(* IEC 61131-3 sources: plcassist-cli/packages/volt-lsp-iec/test-corpus/awa-palletizer/Device/Plc Logic/Application/Library Manager/L_SPMI_PlcParameterManager, 22 files *)

(* ---- L_SPMI_CONSTANT_DEFINES.gvl ---- *)
VAR_GLOBAL
	APPLICATION_AREA_0 : DINT := 0;
	APPLICATION_AREA_1 : DINT := 1;
	APPLICATION_AREA_2 : DINT := 2;
	APPLICATION_AREA_3 : DINT := 3;
END_VAR

(* ---- L_SPMI_LEM_ACCESS.gvl ---- *)
VAR_GLOBAL
	BASIC_SETTINGS : UINT := 4;
	REFID_PLCPM : UINT := 16#2801;
	EVTID_INF_INIT_WRITE : UINT := 16#1101;
	EVTID_INF_DEFAULT_WRITE : UINT := 16#1102;
	EVTID_WRN_INIT_PARAMETER : UINT := 16#1201;
	EVTID_WRN_LOAD_FACTORYSETTINGS : UINT := 16#1202;
	EVTID_WRN_LOAD_TADEFAULTS : UINT := 16#1203;
	EVTID_ERR_REGISTRATION : UINT := 16#1401;
	EVTID_ERR_OPEN_LXD_FILE : UINT := 16#1402;
	EVTID_ERR_OPEN_PRM_FILE : UINT := 16#1403;
	EVTPAR_DT_BOOL : INT := 1;
	EVTPAR_DT_S8 : INT := 2;
	EVTPAR_DT_S16 : INT := 3;
	EVTPAR_DT_S32 : INT := 4;
	EVTPAR_DT_U8 : INT := 5;
	EVTPAR_DT_U16 : INT := 6;
	EVTPAR_DT_U32 : INT := 7;
	EVTPAR_DT_STR_UNI_CODE8 : INT := 8;
	EVTPAR_DT_STR_ASCII : INT := 9;
	EVTPAR_DT_BYTE_ARRAY : INT := 10;
	EVTPAR_DT_S64 : INT := 11;
	EVTPAR_DT_U64 : INT := 12;
	EVTPAR_DT_FLOAT_32 : INT := 13;
	EVTPAR_DT_FLOAT_64 : INT := 14;
END_VAR

(* ---- L_SPMI_ITF_PLCPARAMETERMANAGER.itf ---- *)
INTERFACE L_SPMI_ITF_PLCPARAMETERMANAGER
END_INTERFACE

METHOD GETPARAMETEROBJECT : POINTER TO L_SPMI_ParameterObject
VAR_INPUT
	WINDEX : WORD;
	BYSUBINDEX : BYTE;
	PNUMSUBOBJECTS : POINTER TO BYTE;
END_VAR
END_METHOD

METHOD GETPARAMETEROBJECTLIST : L_SPMI_ParameterObjectList
END_METHOD

METHOD GETPARAMETERVALUE : RTS_IEC_RESULT
VAR_INPUT
	PARAMETERADDRESS : L_SPMI_ParameterAddress;
	PPARAMETERVALUE : POINTER TO L_SPMI_ParameterValueInfo;
END_VAR
END_METHOD

METHOD GETSUBOBJECTRECORDINFO : L_SPMI_SubObjectRecordInfo
VAR_INPUT
	WINDEX : WORD;
END_VAR
END_METHOD

METHOD LOADFACTORYSETTINGS : RTS_IEC_RESULT
END_METHOD

METHOD LOADPARAMETERSET : RTS_IEC_RESULT
END_METHOD

METHOD LOADTADEFAULTPARAMETER : RTS_IEC_RESULT
END_METHOD

METHOD RELAODPARAMETERDESCRIPTION : RTS_IEC_RESULT
END_METHOD

METHOD SAVEPARAMETERSET : RTS_IEC_RESULT
END_METHOD

METHOD SETPARAMETERVALUE : RTS_IEC_RESULT
VAR_INPUT
	PARAMETERADDRESS : L_SPMI_ParameterAddress;
	PPARAMETERVALUE : POINTER TO L_SPMI_ParameterValueInfo;
END_VAR
END_METHOD

METHOD UPDATEONLINECHANGEDPARAMETER : RTS_IEC_RESULT
END_METHOD

(* ---- L_SPMI_UTITF_PLCPM.itf ---- *)
INTERFACE L_SPMI_UTITF_PLCPM
END_INTERFACE

METHOD UT_WRITEPARAMETERVALUE : RTS_IEC_RESULT
VAR_INPUT
	PPARAMETEROBJECT : POINTER TO L_SPMI_ParameterObject;
	PPARAMETERVALUE : POINTER TO L_SPMI_ParameterValueInfo;
	BISDEFAULT : BOOL;
END_VAR
END_METHOD

(* ---- GETBOOLEANPROPERTY.fun ---- *)
FUNCTION GETBOOLEANPROPERTY : BOOL
VAR_INPUT
	STKEY : WSTRING;
END_VAR
END_FUNCTION

(* ---- GETCOMPANY.fun ---- *)
FUNCTION GETCOMPANY : WSTRING
END_FUNCTION

(* ---- GETNUMBERPROPERTY.fun ---- *)
FUNCTION GETNUMBERPROPERTY : DINT
VAR_INPUT
	STKEY : WSTRING;
END_VAR
END_FUNCTION

(* ---- GETTEXTPROPERTY.fun ---- *)
FUNCTION GETTEXTPROPERTY : WSTRING
VAR_INPUT
	STKEY : WSTRING;
END_VAR
END_FUNCTION

(* ---- GETTEXTPROPERTY2.fun ---- *)
FUNCTION GETTEXTPROPERTY2 : POINTER TO WSTRING
VAR_INPUT
	STKEY : WSTRING;
END_VAR
END_FUNCTION

(* ---- GETTITLE.fun ---- *)
FUNCTION GETTITLE : WSTRING
END_FUNCTION

(* ---- GETVERSION.fun ---- *)
FUNCTION GETVERSION : VERSION
END_FUNCTION

(* ---- GETVERSIONPROPERTY.fun ---- *)
FUNCTION GETVERSIONPROPERTY : VERSION
VAR_INPUT
	STKEY : WSTRING;
END_VAR
END_FUNCTION

(* ---- L_SPMI_CONNECTACCESSINTERFACE.fun ---- *)
FUNCTION L_SPMI_CONNECTACCESSINTERFACE : RTS_IEC_RESULT
VAR_INPUT
	PFITERFACE : POINTER TO BYTE;
	ITFTYPE : L_SPMI_InterfaceType;
END_VAR
END_FUNCTION

(* ---- L_SPMI_DISCONNECTACCESSINTERFACE.fun ---- *)
FUNCTION L_SPMI_DISCONNECTACCESSINTERFACE : RTS_IEC_RESULT
VAR_INPUT
	ITFTYPE : L_SPMI_InterfaceType;
END_VAR
END_FUNCTION

(* ---- L_SPMI_READBASEPARAMETER.fun ---- *)
FUNCTION L_SPMI_READBASEPARAMETER : RTS_IEC_RESULT
VAR_INPUT
	WINDEX : WORD;
	BYSUBINDEX : BYTE;
	PPARAMETERVALUE : POINTER TO L_SPMI_ParameterValueInfo;
END_VAR
END_FUNCTION

(* ---- L_SPMI_READBPBPARAMETER.fun ---- *)
FUNCTION L_SPMI_READBPBPARAMETER : RTS_IEC_RESULT
VAR_INPUT
	WINDEX : WORD;
	BYSUBINDEX : BYTE;
	PPARAMETERVALUE : POINTER TO L_SPMI_ParameterValueInfo;
END_VAR
END_FUNCTION

(* ---- L_SPMI_SETPARAMETERMANAGERINSTANCE.fun ---- *)
FUNCTION L_SPMI_SETPARAMETERMANAGERINSTANCE : BOOL
VAR_INPUT
	PPMINSTANCE : POINTER TO BYTE;
END_VAR
END_FUNCTION

(* ---- L_SPMI_WRITEBASEPARAMETER.fun ---- *)
FUNCTION L_SPMI_WRITEBASEPARAMETER : RTS_IEC_RESULT
VAR_INPUT
	WINDEX : WORD;
	BYSUBINDEX : BYTE;
	UISIZE : UINT;
	PPARAMVALUE : POINTER TO BYTE;
END_VAR
END_FUNCTION

(* ---- L_SPMI_WRITEBASEPARAMETER_2.fun ---- *)
FUNCTION L_SPMI_WRITEBASEPARAMETER_2 : RTS_IEC_RESULT
VAR_INPUT
	WINDEX : WORD;
	BYSUBINDEX : BYTE;
	UISIZE : UINT;
	TDATATYPE : L_SPMI_DataType;
	PPARAMVALUE : POINTER TO BYTE;
END_VAR
END_FUNCTION

(* ---- L_SPMI_WRITEBPBPARAMETER.fun ---- *)
FUNCTION L_SPMI_WRITEBPBPARAMETER : RTS_IEC_RESULT
VAR_INPUT
	WINDEX : WORD;
	BYSUBINDEX : BYTE;
	UISIZE : UINT;
	TDATATYPE : L_SPMI_DataType;
	PPARAMVALUE : POINTER TO BYTE;
END_VAR
END_FUNCTION

(* ---- L_SPMI_CRC32.fb ---- *)
FUNCTION_BLOCK L_SPMI_CRC32
VAR
	S_DWCRC32TABLE : ARRAY [0..255] OF DWORD := [16#0, 16#77073096, 16#EE0E612C, 16#990951BA, 16#76DC419, 16#706AF48F, 16#E963A535, 16#9E6495A3, 16#EDB8832, 16#79DCB8A4, 16#E0D5E91E, 16#97D2D988, 16#9B64C2B, 16#7EB17CBD, 16#E7B82D07, 16#90BF1D91, 16#1DB71064, 16#6AB020F2, 16#F3B97148, 16#84BE41DE, 16#1ADAD47D, 16#6DDDE4EB, 16#F4D4B551, 16#83D385C7, 16#136C9856, 16#646BA8C0, 16#FD62F97A, 16#8A65C9EC, 16#14015C4F, 16#63066CD9, 16#FA0F3D63, 16#8D080DF5, 16#3B6E20C8, 16#4C69105E, 16#D56041E4, 16#A2677172, 16#3C03E4D1, 16#4B04D447, 16#D20D85FD, 16#A50AB56B, 16#35B5A8FA, 16#42B2986C, 16#DBBBC9D6, 16#ACBCF940, 16#32D86CE3, 16#45DF5C75, 16#DCD60DCF, 16#ABD13D59, 16#26D930AC, 16#51DE003A, 16#C8D75180, 16#BFD06116, 16#21B4F4B5, 16#56B3C423, 16#CFBA9599, 16#B8BDA50F, 16#2802B89E, 16#5F058808, 16#C60CD9B2, 16#B10BE924, 16#2F6F7C87, 16#58684C11, 16#C1611DAB, 16#B6662D3D, 16#76DC4190, 16#1DB7106, 16#98D220BC, 16#EFD5102A, 16#71B18589, 16#6B6B51F, 16#9FBFE4A5, 16#E8B8D433, 16#7807C9A2, 16#F00F934, 16#9609A88E, 16#E10E9818, 16#7F6A0DBB, 16#86D3D2D, 16#91646C97, 16#E6635C01, 16#6B6B51F4, 16#1C6C6162, 16#856530D8, 16#F262004E, 16#6C0695ED, 16#1B01A57B, 16#8208F4C1, 16#F50FC457, 16#65B0D9C6, 16#12B7E950, 16#8BBEB8EA, 16#FCB9887C, 16#62DD1DDF, 16#15DA2D49, 16#8CD37CF3, 16#FBD44C65, 16#4DB26158, 16#3AB551CE, 16#A3BC0074, 16#D4BB30E2, 16#4ADFA541, 16#3DD895D7, 16#A4D1C46D, 16#D3D6F4FB, 16#4369E96A, 16#346ED9FC, 16#AD678846, 16#DA60B8D0, 16#44042D73, 16#33031DE5, 16#AA0A4C5F, 16#DD0D7CC9, 16#5005713C, 16#270241AA, 16#BE0B1010, 16#C90C2086, 16#5768B525, 16#206F85B3, 16#B966D409, 16#CE61E49F, 16#5EDEF90E, 16#29D9C998, 16#B0D09822, 16#C7D7A8B4, 16#59B33D17, 16#2EB40D81, 16#B7BD5C3B, 16#C0BA6CAD, 16#EDB88320, 16#9ABFB3B6, 16#3B6E20C, 16#74B1D29A, 16#EAD54739, 16#9DD277AF, 16#4DB2615, 16#73DC1683, 16#E3630B12, 16#94643B84, 16#D6D6A3E, 16#7A6A5AA8, 16#E40ECF0B, 16#9309FF9D, 16#A00AE27, 16#7D079EB1, 16#F00F9344, 16#8708A3D2, 16#1E01F268, 16#6906C2FE, 16#F762575D, 16#806567CB, 16#196C3671, 16#6E6B06E7, 16#FED41B76, 16#89D32BE0, 16#10DA7A5A, 16#67DD4ACC, 16#F9B9DF6F, 16#8EBEEFF9, 16#17B7BE43, 16#60B08ED5, 16#D6D6A3E8, 16#A1D1937E, 16#38D8C2C4, 16#4FDFF252, 16#D1BB67F1, 16#A6BC5767, 16#3FB506DD, 16#48B2364B, 16#D80D2BDA, 16#AF0A1B4C, 16#36034AF6, 16#41047A60, 16#DF60EFC3, 16#A867DF55, 16#316E8EEF, 16#4669BE79, 16#CB61B38C, 16#BC66831A, 16#256FD2A0, 16#5268E236, 16#CC0C7795, 16#BB0B4703, 16#220216B9, 16#5505262F, 16#C5BA3BBE, 16#B2BD0B28, 16#2BB45A92, 16#5CB36A04, 16#C2D7FFA7, 16#B5D0CF31, 16#2CD99E8B, 16#5BDEAE1D, 16#9B64C2B0, 16#EC63F226, 16#756AA39C, 16#26D930A, 16#9C0906A9, 16#EB0E363F, 16#72076785, 16#5005713, 16#95BF4A82, 16#E2B87A14, 16#7BB12BAE, 16#CB61B38, 16#92D28E9B, 16#E5D5BE0D, 16#7CDCEFB7, 16#BDBDF21, 16#86D3D2D4, 16#F1D4E242, 16#68DDB3F8, 16#1FDA836E, 16#81BE16CD, 16#F6B9265B, 16#6FB077E1, 16#18B74777, 16#88085AE6, 16#FF0F6A70, 16#66063BCA, 16#11010B5C, 16#8F659EFF, 16#F862AE69, 16#616BFFD3, 16#166CCF45, 16#A00AE278, 16#D70DD2EE, 16#4E048354, 16#3903B3C2, 16#A7672661, 16#D06016F7, 16#4969474D, 16#3E6E77DB, 16#AED16A4A, 16#D9D65ADC, 16#40DF0B66, 16#37D83BF0, 16#A9BCAE53, 16#DEBB9EC5, 16#47B2CF7F, 16#30B5FFE9, 16#BDBDF21C, 16#CABAC28A, 16#53B39330, 16#24B4A3A6, 16#BAD03605, 16#CDD70693, 16#54DE5729, 16#23D967BF, 16#B3667A2E, 16#C4614AB8, 16#5D681B02, 16#2A6F2B94, 16#B40BBE37, 16#C30C8EA1, 16#5A05DF1B, 16#2D02EF8D];
END_VAR
END_FUNCTION_BLOCK

METHOD UPDATECRC : DWORD
VAR_INPUT
	DWCRC : DWORD;
	PDATA : POINTER TO BYTE;
	DWSIZE : __XWORD;
END_VAR
END_METHOD

(* ---- L_SPMI_PLCPARAMETERMANAGER.fb ---- *)
FUNCTION_BLOCK L_SPMI_PLCPARAMETERMANAGER
VAR
	M_SZAPPNAME2 : STRING;
	M_DWPARAMOBJVERSION : DWORD;
	M_BUNITTEST : BOOL := FALSE;
	FBINIT : BOOL;
	FBAFTERGLOBALINIT : BOOL;
	XLXDFILENOTEXIST : BOOL;
	XPRMFILENOTEXIST : BOOL;
	M_UICNTALLMEM : UINT;
	M_UICNTPERSISTMEM : UINT;
	M_UICNTSTORE : UINT;
	M_UINOTCNTSTORE : UINT;
	M_UICNTPLCSTORE : UINT;
	M_BSTOREDONE : BOOL;
	M_BOOTPROJPATH : STRING;
	M_SZCMPNAME : STRING := 'PLC_PM';
	M_BLXDLOADED : BOOL;
	M_PPARAMOBJECTMEM : POINTER TO BYTE;
	M_PSINGLEPARAMOBJECTSMEM : POINTER TO BYTE;
	M_PCUROBJLISTELEMENT : POINTER TO L_SPMI_ObjectList;
	M_PCURPARAMETEROBJECT : POINTER TO L_SPMI_ParameterObject;
	M_PCURSINGLEPARAMETEROBJECT : POINTER TO L_SPMI_ParameterObject;
	M_DWNUMBEROFOBJECTS : DWORD := 0;
	M_PFIRSTPARAMETEROBJECT : POINTER TO L_SPMI_ParameterObject := 0;
	M_PPREVPARAMETEROBJECT : POINTER TO L_SPMI_ParameterObject := 0;
	M_POBJECTTEMPLATELIST : POINTER TO BYTE := 0;
	M_PCUROBJECTTEMPLATE : POINTER TO L_SPMI_ObjectTemplate := 0;
	M_UICOUNTOBJECTTEMPLATES : UINT := 0;
	M_BISOBJECTTEMPLATE : BOOL := FALSE;
	M_BSUBOBJRECORD : BOOL;
	M_BSINGLEOBJECTPARAM : BOOL;
	M_BOVERWRITTENBASEPARAM : BOOL;
	M_PFIRSTPERSISTENTPARAM : POINTER TO L_SPMI_ParameterObject;
	M_PPREVPERSISTENTPARAM : POINTER TO L_SPMI_ParameterObject;
	M_UITADEFAULTNUMBER : UINT;
	M_BPARAMETERGROUPTADEFAULT : BOOL;
	M_PFIRSTTADEFAULTPARAMETER : POINTER TO L_SPMI_ParameterObject;
	M_PPREVTADEFAULTPARAMETER : POINTER TO L_SPMI_ParameterObject;
	M_PFIRSTBASETADEFAULTPARAMETER : POINTER TO L_SPMI_ParameterObject;
	M_PPREVBASETADEFAULTPARAMETER : POINTER TO L_SPMI_ParameterObject;
	M_PBASETADEFAULTPARAMETERLIST : POINTER TO BYTE;
	M_PCURBASETADEFAULTOBJECT : POINTER TO L_SPMI_ParameterObject;
	M_PCURSELECTLISTELEMENT : POINTER TO BYTE;
	M_PATTRLOWLIMIT : POINTER TO STRING(255);
	M_PATTRHIGHLIMIT : POINTER TO STRING(255);
	M_PATTRDEFAULT : POINTER TO STRING(255);
	M_STRLOWLIMIT : STRING(255);
	M_STRHIGHLIMIT : STRING(255);
	M_STRDEFAULTVALUE : STRING(255);
	M_PAPPLICATION : POINTER TO APPLICATION;
	M_SZAPPNAME : STRING(MAX_LEN_APPLNAME);
	M_PAPPDATA : POINTER TO BYTE;
	M_PAPPAREA_0 : POINTER TO BYTE;
	M_PAPPAREA_1 : POINTER TO BYTE;
	M_PAPPAREA_2 : POINTER TO BYTE;
	M_PAPPAREA_3 : POINTER TO BYTE;
	M_CUROBJINDEX : WORD;
	M_UIOBJECTLISTNUMBER : UINT;
	M_BYSUBOBJECTNUMBER : BYTE;
	M_UITEMPLATELISTNUMBER : UINT;
	M_UICOUNTSUBOBJECT : UINT;
	M_FILEHEADER : L_SPMI_FileHeader;
	M_DATAHEADER : L_SPMI_DataHeader;
	M_PPRMDATA : POINTER TO BYTE;
	M_DWPRMDATASIZE : DWORD;
	M_SZPATHLXDFILE : STRING(255);
	M_SZPATHPRMFILE : STRING(255);
	M_SZPATHALLACTPARAMS : STRING(255);
	M_SZPATHPRMFILE_TEMP : STRING(255);
	M_SZPATHPRMFILE_TEST : STRING(255);
	M_SZPATHPRMFILE_PRG : STRING(255);
	M_SZPATHUPDATEONLINECHANGEDPARAMETER : STRING(255);
	M_SZPATHUPDATEONLINECHANGEDPARAMETERTRIGGERINSIMULATIONMODE : STRING(255);
	M_ABYPRMBUFFER : ARRAY [0..999] OF BYTE;
	M_ABYZEROBUFFER : ARRAY [0..255] OF BYTE;
	M_HEVENTPARVALUECHANGED : RTS_IEC_HANDLE;
	M_EVENTPARAM_VALCHANGED : CmpEventMgr.EventParam;
	M_PARAVALUECHANGED : L_SSYP.L_SSYP_EVTPARAM_CmpLenzeIPCSystemSoftPLCParaChanged;
	M_HEVENTPARDESCRIPTIONLOADED : RTS_IEC_HANDLE;
	M_EVENTPARAM_PARDESCLOADED : CmpEventMgr.EventParam;
	M_HEVENTDOWNLOADDONE : RTS_IEC_HANDLE;
	M_HEVENTRESETDONE : RTS_IEC_HANDLE;
	M_HEVENTCOMMCYCLEINSIMULATIONMODE : RTS_IEC_HANDLE;
	M_HINTERFACEDOWNLOADDONE : RTS_IEC_HANDLE;
	M_HINTERFACERESETDONE : RTS_IEC_HANDLE;
	M_HINTERFACECOMMCYCLEINSIMULATIONMODE : RTS_IEC_HANDLE;
	M_HEVENTUPDATECONFIGURATIONDONE : RTS_IEC_HANDLE;
	M_HINTERFACEUPDATECONFIGURATIONDONE : RTS_IEC_HANDLE;
	M_ITFEVENTCALLBACK : CmpEventMgr.ICmpEventCallback;
	M_TASKHANDLE : RTS_IEC_HANDLE;
	M_CURTASKPRIO : UDINT;
	FBCRC32 : L_SPMI_CRC32;
	M_HTRACEFILE : RTS_IEC_HANDLE;
	M_SZPATHTRACEFILE : STRING;
	M_SZPATHTRACEFILE_RENAME : STRING;
	M_SZNEWLINE : STRING := '$N';
	M_EERRSTOREPRM : UINT;
	M_UISTORE : UINT;
	M_BLXDFILEREAD : BOOL := FALSE;
	M_BOBJECTLISTLOADED : BOOL := FALSE;
	M_UIPARAMETERCOUNT : UINT := 0;
	M_HLENZEMODULEHANDLER : RTS_IEC_HANDLE := 0;
	M_HLENZEERRORMANAGER : RTS_IEC_HANDLE := 0;
	M_SZTRACETEXT : STRING;
	M_RESULT : RTS_IEC_RESULT;
	M_TONCHECKONLINECHANGEPARAFILE : TON;
	SINSTANCESTRFULL : STRING(255);
	LXDFILEREAD : BOOL;
	OBJECTLISTLOADED : BOOL;
	OBJECTLISTNUMBER : UINT;
	PARAMETERGROUPTADEFAULTSLOADED : BOOL;
	PARAMETEROBJECTSCOUNT : UINT;
END_VAR
END_FUNCTION_BLOCK

METHOD EVENTCALLBACK : UDINT
VAR_INPUT
	PEVENTPARAM : POINTER TO EventParam;
END_VAR
END_METHOD

METHOD FB_AFTERGLOABALINIT : BOOL
END_METHOD

METHOD FB_EXIT : BOOL
VAR_INPUT
	BINCOPYCODE : BOOL;
END_VAR
END_METHOD

METHOD FB_INIT : BOOL
VAR_INPUT
	BINITRETAINS : BOOL;
	BINCOPYCODE : BOOL;
END_VAR
END_METHOD

METHOD GETSUBOBJCOUNT_X : UINT
END_METHOD

METHOD CHECKVALUELIMITS_1_X : RTS_IEC_RESULT
VAR_INPUT
	PARAMETERVALUE : L_SPMI_ParameterValueInfo;
	PPARAMVALUELIMITS : POINTER TO L_SPMI_Limits;
END_VAR
END_METHOD

METHOD CHECKVALUELIMITS_2_X : RTS_IEC_RESULT
VAR_INPUT
	PARAMETERVALUE : L_SPMI_ParameterValueInfo;
	PPARAMVALUELIMITS : POINTER TO L_SPMI_Limits;
	DATATYPE : L_SPMI_DataType;
END_VAR
END_METHOD

METHOD INITIALIZEPRMDATA_1_X : RTS_IEC_RESULT
VAR_INPUT
	PDATAHEADER : POINTER TO L_SPMI_DataHeader;
	PPRMDATA : POINTER TO BYTE;
END_VAR
END_METHOD

METHOD INITIALIZEPRMDATA_X : RTS_IEC_RESULT
VAR_INPUT
	PDATAHEADER : POINTER TO L_SPMI_DataHeader;
	PPRMDATA : POINTER TO BYTE;
END_VAR
END_METHOD

METHOD SCALEEXTERNTOINTERNVALUE_1_X : RTS_IEC_RESULT
VAR_INPUT
	PEXTERNVAL : POINTER TO L_SPMI_ParameterValueInfo;
	PINTERNVAL : POINTER TO BYTE;
	PINTERNVALSIZE : POINTER TO UINT;
	PPARAMOBJ : POINTER TO L_SPMI_ParameterObject;
END_VAR
END_METHOD

METHOD STOREPRMFILE_1_X : RTS_IEC_RESULT
END_METHOD

METHOD STOREPRMFILE_X : RTS_IEC_RESULT
END_METHOD

METHOD UPDATEPARSETCFG_X : RTS_IEC_RESULT
VAR_INPUT
	SZPRMFILENAME : STRING;
	NEWPRMFILECRC : DWORD;
END_VAR
END_METHOD

METHOD WRITEPARAMETERVALUE_1_X : RTS_IEC_RESULT
VAR_INPUT
	PPARAMOBJ : POINTER TO L_SPMI_ParameterObject;
	PPARAMETERVALUE : POINTER TO L_SPMI_ParameterValueInfo;
END_VAR
END_METHOD

METHOD WRITEPARAMETERVALUE_2_X : RTS_IEC_RESULT
VAR_INPUT
	PPARAMOBJ : POINTER TO L_SPMI_ParameterObject;
	PPARAMETERVALUE : POINTER TO L_SPMI_ParameterValueInfo;
END_VAR
END_METHOD

METHOD WRITEPARAMETERVALUE_DEFAULT_X : RTS_IEC_RESULT
VAR_INPUT
	PPARAMOBJ : POINTER TO L_SPMI_ParameterObject;
	PPARAMETERVALUE : POINTER TO L_SPMI_ParameterValueInfo;
END_VAR
END_METHOD

METHOD GETPARAMETEROBJECT : POINTER TO L_SPMI_ParameterObject
VAR_INPUT
	WINDEX : WORD;
	BYSUBINDEX : BYTE;
	PNUMSUBOBJECTS : POINTER TO BYTE;
END_VAR
END_METHOD

METHOD GETPARAMETEROBJECTLIST : L_SPMI_ParameterObjectList
END_METHOD

METHOD GETPARAMETERVALUE : RTS_IEC_RESULT
VAR_INPUT
	PARAMETERADDRESS : L_SPMI_ParameterAddress;
	PPARAMETERVALUE : POINTER TO L_SPMI_ParameterValueInfo;
END_VAR
END_METHOD

METHOD GETSUBOBJECTRECORDINFO : L_SPMI_SubObjectRecordInfo
VAR_INPUT
	WINDEX : WORD;
END_VAR
END_METHOD

METHOD LOADFACTORYSETTINGS : RTS_IEC_RESULT
END_METHOD

METHOD LOADPARAMETERSET : RTS_IEC_RESULT
END_METHOD

METHOD LOADTADEFAULTPARAMETER : RTS_IEC_RESULT
END_METHOD

METHOD RELAODPARAMETERDESCRIPTION : RTS_IEC_RESULT
END_METHOD

METHOD SAVEALLACTUALPARAMS : RTS_IEC_RESULT
END_METHOD

METHOD SAVEPARAMETERSET : RTS_IEC_RESULT
END_METHOD

METHOD SETPARAMETERVALUE : RTS_IEC_RESULT
VAR_INPUT
	PARAMETERADDRESS : L_SPMI_ParameterAddress;
	PPARAMETERVALUE : POINTER TO L_SPMI_ParameterValueInfo;
END_VAR
END_METHOD

METHOD UPDATEONLINECHANGEDPARAMETER : RTS_IEC_RESULT
END_METHOD

METHOD INITIALIZEALLPARAMETER : RTS_IEC_RESULT
END_METHOD

METHOD INITIALIZEBPBPARAMETER : RTS_IEC_RESULT
END_METHOD

METHOD INITIALIZEPLCPARAMETER : RTS_IEC_RESULT
END_METHOD

METHOD SENDALLVALUECHANGEDEVENTS : RTS_IEC_RESULT
END_METHOD

METHOD GETPOINTERTOPARAMETERVALUE : L_SPMI_PointerToValue
VAR_INPUT
	WINDEX : WORD;
	BYSUBINDEX : BYTE;
END_VAR
END_METHOD

METHOD ANALYZETAG : RTS_IEC_RESULT
VAR_INPUT
	PTAGINFO : POINTER TO L_SPMI_TagInformation;
END_VAR
END_METHOD

METHOD FINDCLOSETAG : RTS_IEC_RESULT
VAR_INPUT
	PTAGINFO : POINTER TO L_SPMI_TagInformation;
	PENDBUFFER : POINTER TO BYTE;
END_VAR
END_METHOD

METHOD FINDOPENTAG : RTS_IEC_RESULT
VAR_INPUT
	PTAGINFO : POINTER TO L_SPMI_TagInformation;
	PSTARTPOS : POINTER TO BYTE;
	PENDBUFFER : POINTER TO BYTE;
END_VAR
END_METHOD

METHOD GETATTRIBUTEVALUE : POINTER TO STRING
VAR_INPUT
	PELEMENTINFO : POINTER TO L_SPMI_ElementInfo;
	SZATTRIBUTENAME : STRING;
END_VAR
END_METHOD

METHOD GETELEMENT : RTS_IEC_RESULT
VAR_INPUT
	PCURBYTE : POINTER TO BYTE;
	PELEMENTINFO : POINTER TO L_SPMI_ElementInfo;
END_VAR
END_METHOD

METHOD GETTAGINFO : RTS_IEC_RESULT
VAR_INPUT
	PTAGINFO : POINTER TO L_SPMI_TagInformation;
END_VAR
END_METHOD

METHOD PARSELXDFILE : RTS_IEC_RESULT
VAR_INPUT
	SZFILE : REFERENCE TO STRING;
END_VAR
END_METHOD

METHOD READPARAMETERVALUE : RTS_IEC_RESULT
VAR_INPUT
	PPARAMOBJ : POINTER TO L_SPMI_ParameterObject;
	PPARAMETERVALUE : POINTER TO L_SPMI_ParameterValueInfo;
END_VAR
END_METHOD

METHOD WRITEPARAMETERVALUE : RTS_IEC_RESULT
VAR_INPUT
	PPARAMETEROBJECT : POINTER TO L_SPMI_ParameterObject;
	PPARAMETERVALUE : POINTER TO L_SPMI_ParameterValueInfo;
	BISDEFAULT : BOOL;
END_VAR
END_METHOD

METHOD WRITEPRMDATAONLINECHANGED : RTS_IEC_RESULT
VAR_INPUT
	PDATAHEADER : POINTER TO L_SPMI_DataHeader;
	PPRMDATA : POINTER TO BYTE;
END_VAR
END_METHOD

METHOD STOREPARSETCONFIG
VAR_INPUT
	DWPRMCRC : DWORD;
END_VAR
END_METHOD

METHOD STOREPRMFILE_BASE_AND_PLC : RTS_IEC_RESULT
END_METHOD

METHOD STOREPRMFILE_ONLY_PLC : RTS_IEC_RESULT
END_METHOD

METHOD STOREPRMFILE_OVERWRITEBASE_AND_STOREPLC : RTS_IEC_RESULT
END_METHOD

METHOD WRITEZEROBUFFERTOFILE : RTS_IEC_RESULT
VAR_INPUT
	HFILE : RTS_IEC_HANDLE;
	DWSIZE : DWORD;
END_VAR
END_METHOD

METHOD UT_WRITEPARAMETERVALUE : RTS_IEC_RESULT
VAR_INPUT
	PPARAMETEROBJECT : POINTER TO L_SPMI_ParameterObject;
	PPARAMETERVALUE : POINTER TO L_SPMI_ParameterValueInfo;
	BISDEFAULT : BOOL;
END_VAR
END_METHOD

METHOD CLEANLXDDATA : RTS_IEC_RESULT
END_METHOD

METHOD CLEANPRMDATA : RTS_IEC_RESULT
END_METHOD

METHOD FREEALLOCATEDMEM
END_METHOD

METHOD GETAPPAREA : POINTER TO BYTE
VAR_INPUT
	UIAREA : UINT;
END_VAR
END_METHOD

METHOD GETOVERWRITTENPARAMOBJ : POINTER TO L_SPMI_ParameterObject
VAR_INPUT
	WINDEX : WORD;
	BYSUBINDEX : BYTE;
END_VAR
END_METHOD

METHOD GETPARAMOBJ : POINTER TO L_SPMI_ParameterObject
VAR_INPUT
	WINDEX : WORD;
	BYSUBINDEX : BYTE;
	PNUMSUBOBJECTS : POINTER TO BYTE;
	PRESULT : POINTER TO RTS_IEC_RESULT;
END_VAR
END_METHOD

METHOD GETPERSISTENTPARAMOBJ : POINTER TO L_SPMI_ParameterObject
VAR_INPUT
	WINDEX : WORD;
	BYSUBINDEX : BYTE;
END_VAR
END_METHOD

METHOD LOADLXDDATA : RTS_IEC_RESULT
VAR_INPUT
	SZFILE : REFERENCE TO STRING;
END_VAR
END_METHOD

METHOD LOADPRMDATA : POINTER TO BYTE
VAR_INPUT
	SZFILE : REFERENCE TO STRING;
	PFILEHEADER : POINTER TO L_SPMI_FileHeader;
	PDATAHEADER : POINTER TO L_SPMI_DataHeader;
END_VAR
END_METHOD

METHOD GETPRMPARAMETER : POINTER TO L_SPMI_ParameterHeader
VAR_INPUT
	WINDEX : WORD;
	BYSUBINDEX : BYTE;
	PLASTPARAMHEADER : POINTER TO L_SPMI_ParameterHeader;
END_VAR
END_METHOD

METHOD GETPRMVALUE : RTS_IEC_RESULT
VAR_INPUT
	PPARAMDATA : POINTER TO BYTE;
	PPARAMHEADER : POINTER TO L_SPMI_ParameterHeader;
	PPARAMOBJ : POINTER TO L_SPMI_ParameterObject;
	PPARAMVALUE : POINTER TO L_SPMI_ParameterValue;
END_VAR
END_METHOD

METHOD GETDATATYPE : L_SPMI_DataType
VAR_INPUT
	PSTRINGVALUE : POINTER TO STRING;
END_VAR
END_METHOD

METHOD GETPARAMETERTYPE : L_SPMI_ParameterType
VAR_INPUT
	PSTRINGVALUE : POINTER TO STRING;
END_VAR
END_METHOD

METHOD INITPARAMETEROBJECT
VAR_INPUT
	PPARAMOBJECT : POINTER TO L_SPMI_ParameterObject;
END_VAR
END_METHOD

METHOD SETDATASIZE : RTS_IEC_RESULT
VAR_INPUT
	PPARAMETEROBJECT : POINTER TO L_SPMI_ParameterObject;
END_VAR
END_METHOD

METHOD SETDEFAULTVALUE : RTS_IEC_RESULT
VAR_INPUT
	PPARAMETEROBJECT : POINTER TO L_SPMI_ParameterObject;
	PVALUEASSTRING : POINTER TO STRING(255);
END_VAR
END_METHOD

METHOD SETREFTEMPLATE
VAR_INPUT
	PPARAMETEROBJECT : POINTER TO L_SPMI_ParameterObject;
	PTEMPLATENAME : POINTER TO STRING;
END_VAR
END_METHOD

METHOD SETSELECTTEXTVALUE : RTS_IEC_RESULT
VAR_INPUT
	PSELECTTEXTVALUE : POINTER TO BYTE;
	PVALUEASSTRING : POINTER TO STRING;
	DATATYPE : L_SPMI_DataType;
END_VAR
END_METHOD

METHOD SETVALUELIMITS : RTS_IEC_RESULT
VAR_INPUT
	PPARAMETEROBJECT : POINTER TO L_SPMI_ParameterObject;
	PLOWLIMITASSTRING : POINTER TO STRING;
	PHIGHLIMITASSTRING : POINTER TO STRING;
END_VAR
END_METHOD

METHOD CHECKSELECTLIST : RTS_IEC_RESULT
VAR_INPUT
	PPARAMVALUE : POINTER TO L_SPMI_ParameterValue;
	PPARAMSELECTLIST : POINTER TO L_SPMI_SelectList;
END_VAR
END_METHOD

METHOD CHECKSELECTLIST_1 : RTS_IEC_RESULT
VAR_INPUT
	PARAMETERVALUE : L_SPMI_ParameterValueInfo;
	PPARAMSELECTLIST : POINTER TO L_SPMI_SelectList;
END_VAR
END_METHOD

METHOD CHECKVALUELIMITS : RTS_IEC_RESULT
VAR_INPUT
	PPARAMVALUE : POINTER TO L_SPMI_ParameterValue;
	PPARAMVALUELIMITS : POINTER TO L_SPMI_Limits;
END_VAR
END_METHOD

METHOD CHECKVALUESIZE : RTS_IEC_RESULT
VAR_INPUT
	UIDATASIZE : UINT;
	PPARAMOBJ : POINTER TO L_SPMI_ParameterObject;
END_VAR
END_METHOD

METHOD ISPERSISTENPLCPARAMETER : BOOL
VAR_INPUT
	WINDEX : WORD;
	BYSUBINDEX : BYTE;
END_VAR
END_METHOD

METHOD SCALEEXTERNTOINTERNVALUE : RTS_IEC_RESULT
VAR_INPUT
	PEXTERNVAL : POINTER TO L_SPMI_ParameterValueInfo;
	PINTERNVAL : POINTER TO BYTE;
	PPARAMOBJ : POINTER TO L_SPMI_ParameterObject;
END_VAR
END_METHOD

METHOD SCALEEXTERNTOINTERNVALUE_2 : RTS_IEC_RESULT
VAR_INPUT
	PEXTERNVAL : POINTER TO L_SPMI_ParameterValueInfo;
	PINTERNVAL : POINTER TO L_SPMI_ParameterValue;
	PPARAMOBJ : POINTER TO L_SPMI_ParameterObject;
END_VAR
END_METHOD

METHOD SCALEINTERNTOEXTERNVALUE : RTS_IEC_RESULT
VAR_INPUT
	PINTERNVAL : POINTER TO BYTE;
	PPARAMETERVALUE : POINTER TO L_SPMI_ParameterValueInfo;
	PPARAMOBJ : POINTER TO L_SPMI_ParameterObject;
END_VAR
END_METHOD
